(* IEC 61131-3 sources: PLCHoney/Boston Intersection Models/plc_template/webserver/example_st_files, 7 files *)

(* ---- BACNet.st ---- *)
FUNCTION_BLOCK Simulator
  VAR_OUTPUT
    Out : REAL;
  END_VAR
  VAR_INPUT
    MinVal : REAL;
    MaxVal : REAL;
    PeriodSeconds : INT;
  END_VAR
  VAR
    TON0 : TON;
    seconds : INT;
    BaseVal : REAL;
    VarVal : REAL;
  END_VAR

  (* pseudo-random variations *)
  TON0(IN := TRUE, PT := T#3120s);
  IF TON0.Q THEN
    TON0(IN := FALSE);
  END_IF;
  seconds := TIME_TO_INT(TON0.ET);

  BaseVal := (MaxVal + MinVal)/2.0;
  VarVal  := (MaxVal-MinVal)*INT_TO_REAL((seconds MOD PeriodSeconds) - (PeriodSeconds/2))/INT_TO_REAL(PeriodSeconds);

  Out :=  BaseVal + VarVal;
END_FUNCTION_BLOCK

PROGRAM program0
  VAR
    EnergyCounter AT %MD0.2.0 : REAL;
    Temperature AT %ID0.0.0 : REAL;
    Humidity AT %ID0.0.1 : REAL;
  END_VAR
  VAR
    TempSimulation : Simulator;
    HumiditySimulation : Simulator;
  END_VAR
  VAR
    TemperatureSetPoint AT %QD0.1.0 : REAL;
    ControlDisable AT %QX0.4.2 : BOOL;
    Heater AT %IX0.3.0 : BOOL;
    Cooler AT %IX0.3.1 : BOOL;
  END_VAR
  VAR
    ADD3_OUT : REAL;
    GT16_OUT : BOOL;
    AND19_OUT : BOOL;
    LT17_OUT : BOOL;
    AND24_OUT : BOOL;
  END_VAR

  ADD3_OUT := ADD(EnergyCounter, 0.00131);
  EnergyCounter := ADD3_OUT;
  TempSimulation(MinVal := 18.0, MaxVal := 30.0, PeriodSeconds := 120);
  Temperature := TempSimulation.Out;
  HumiditySimulation(MinVal := 55.0, MaxVal := 78.0, PeriodSeconds := 58);
  Humidity := HumiditySimulation.Out;
  GT16_OUT := GT(Temperature, TemperatureSetPoint);
  AND19_OUT := AND(NOT(ControlDisable), GT16_OUT);
  Cooler := AND19_OUT;
  LT17_OUT := LT(Temperature, TemperatureSetPoint);
  AND24_OUT := AND(NOT(ControlDisable), LT17_OUT);
  Heater := AND24_OUT;
END_PROGRAM

CONFIGURATION config

  RESOURCE resource1 ON PLC
    TASK task0(INTERVAL := T#20ms,PRIORITY := 0);
    PROGRAM instance0 WITH task0 : program0;
  END_RESOURCE
END_CONFIGURATION

(* ---- First_Steps.st ---- *)
FUNCTION_BLOCK CounterSFC
  VAR_INPUT
    Reset : BOOL;
  END_VAR
  VAR_OUTPUT
    OUT : INT;
  END_VAR
  VAR
    Cnt : INT;
  END_VAR
  VAR_EXTERNAL CONSTANT
    ResetCounterValue : INT;
  END_VAR

  INITIAL_STEP Start:
  END_STEP

  TRANSITION FROM Start TO ResetCounter
    := Reset;
  END_TRANSITION

  STEP ResetCounter:
    RESETCOUNTER_INLINE1(N);
    RESETCOUNTER_INLINE2(N);
  END_STEP

  ACTION RESETCOUNTER_INLINE1:
    Cnt := ResetCounterValue;
  END_ACTION

  ACTION RESETCOUNTER_INLINE2:
    OUT := Cnt;
  END_ACTION

  TRANSITION FROM ResetCounter TO Start
    := NOT Reset;
  END_TRANSITION

  TRANSITION FROM Start TO Count
    := NOT Reset;
  END_TRANSITION

  STEP Count:
    COUNT_INLINE3(N);
    COUNT_INLINE4(N);
  END_STEP

  ACTION COUNT_INLINE3:
    Cnt := Cnt + 1;
  END_ACTION

  ACTION COUNT_INLINE4:
    OUT := Cnt;
  END_ACTION

  TRANSITION FROM Count TO Start
    := Reset;
  END_TRANSITION

END_FUNCTION_BLOCK

FUNCTION_BLOCK CounterFBD
  VAR_INPUT
    Reset : BOOL;
  END_VAR
  VAR_OUTPUT
    OUT : INT;
  END_VAR
  VAR
    Cnt : INT;
  END_VAR
  VAR_EXTERNAL CONSTANT
    ResetCounterValue : INT;
  END_VAR
  VAR
    ADD4_OUT : INT;
    SEL7_OUT : INT;
  END_VAR

  ADD4_OUT := ADD(1, Cnt);
  SEL7_OUT := SEL(Reset, ADD4_OUT, ResetCounterValue);
  Cnt := SEL7_OUT;
  OUT := Cnt;
END_FUNCTION_BLOCK

FUNCTION_BLOCK CounterIL
  VAR
    Cnt : INT;
  END_VAR
  VAR_INPUT
    Reset : BOOL;
  END_VAR
  VAR_OUTPUT
    OUT : INT;
  END_VAR
  VAR_EXTERNAL CONSTANT
    ResetCounterValue : INT;
  END_VAR

  LD Reset
  JMPC ResetCnt

  (* increment counter *)
  LD Cnt
  ADD 1
  JMP QuitFb

  ResetCnt:
  (* reset counter *)
  LD ResetCounterValue

  QuitFb:
  (* save results *)
  ST Cnt
  ST Out
END_FUNCTION_BLOCK

FUNCTION AverageVal : REAL
  VAR_INPUT
    Cnt1 : INT;
    Cnt2 : INT;
    Cnt3 : INT;
    Cnt4 : INT;
    Cnt5 : INT;
  END_VAR
  VAR
    InputsNumber : REAL := 5.0;
  END_VAR

  AverageVal := INT_TO_REAL(Cnt1+Cnt2+Cnt3+Cnt4+Cnt5)/InputsNumber;
END_FUNCTION

FUNCTION_BLOCK CounterST
  VAR_INPUT
    Reset : BOOL;
  END_VAR
  VAR
    Cnt : INT;
  END_VAR
  VAR_OUTPUT
    OUT : INT;
  END_VAR
  VAR_EXTERNAL CONSTANT
    ResetCounterValue : INT;
  END_VAR

  IF Reset THEN
    Cnt := ResetCounterValue;
  ELSE
    Cnt := Cnt + 1;
  END_IF;

  Out := Cnt;
END_FUNCTION_BLOCK

FUNCTION_BLOCK CounterLD
  VAR_INPUT
    Reset : BOOL;
  END_VAR
  VAR_OUTPUT
    Out : INT;
  END_VAR
  VAR
    Cnt : INT;
  END_VAR
  VAR_EXTERNAL CONSTANT
    ResetCounterValue : INT;
  END_VAR
  VAR
    ADD4_OUT : INT;
    SEL7_OUT : INT;
  END_VAR

  ADD4_OUT := ADD(1, Cnt);
  SEL7_OUT := SEL(Reset, ADD4_OUT, ResetCounterValue);
  Cnt := SEL7_OUT;
  Out := Cnt;
END_FUNCTION_BLOCK

PROGRAM plc_prg
  VAR_INPUT
    Reset : BOOL;
  END_VAR
  VAR_OUTPUT
    Cnt1 : INT;
    Cnt2 : INT;
    Cnt3 : INT;
    Cnt4 : INT;
    Cnt5 : INT;
  END_VAR
  VAR
    CounterST0 : CounterST;
    CounterFBD0 : CounterFBD;
    CounterSFC0 : CounterSFC;
    CounterIL0 : CounterIL;
    CounterLD0 : CounterLD;
    AVCnt : REAL;
    AverageVal17_OUT : REAL;
  END_VAR

  CounterST0(Reset := Reset);
  Cnt1 := CounterST0.OUT;
  AverageVal17_OUT := AverageVal(Cnt1, Cnt2, Cnt3, Cnt4, Cnt5);
  AVCnt := AverageVal17_OUT;
  CounterFBD0(Reset := Reset);
  Cnt2 := CounterFBD0.OUT;
  CounterSFC0(Reset := Reset);
  Cnt3 := CounterSFC0.OUT;
  CounterIL0(Reset := Reset);
  Cnt4 := CounterIL0.OUT;
  CounterLD0(Reset := Reset);
  Cnt5 := CounterLD0.Out;
END_PROGRAM

CONFIGURATION config
  VAR_GLOBAL CONSTANT
    ResetCounterValue : INT := 17;
  END_VAR

  RESOURCE resource1 ON PLC
    TASK plc_task(INTERVAL := T#100ms,PRIORITY := 1);
    PROGRAM plc_task_instance WITH plc_task : plc_prg;
  END_RESOURCE
END_CONFIGURATION

(* ---- modbus.st ---- *)
FUNCTION_BLOCK Generator
  VAR_OUTPUT
    OUT : BOOL;
  END_VAR
  VAR_INPUT
    PON : TIME;
    POFF : TIME;
  END_VAR
  VAR
    T1 : TON;
    T2 : TOF;
  END_VAR

  T1( IN := NOT T2.Q, PT := POFF);
  T2( IN := T1.Q,     PT := PON);
  OUT := T2.Q;
END_FUNCTION_BLOCK

PROGRAM program0
  VAR
    Counter : INT;
    CounterReadBack : INT;
  END_VAR
  VAR
    MasterWriteToReg0 AT %QW0.0.0.0 : INT;
    MasterReadFromReg1 AT %IW0.0.1.0 : INT;
    SlaveHoldReg0 AT %IW0.1.0.0 : WORD;
    SlaveInputReg0 AT %QW0.1.1.0 : WORD;
  END_VAR
  VAR
    CTU0 : CTU;
    Generator0 : Generator;
    R_TRIG1 : R_TRIG;
  END_VAR

  Generator0(PON := T#1s, POFF := T#1s);
  R_TRIG1(CLK := Generator0.OUT);
  CTU0(CU := R_TRIG1.Q, PV := 32767);
  Counter := CTU0.CV;
  MasterWriteToReg0 := Counter;
  CounterReadBack := MasterReadFromReg1;
  SlaveInputReg0 := SlaveHoldReg0;
END_PROGRAM

CONFIGURATION config

  RESOURCE resource1 ON PLC
    TASK task0(INTERVAL := T#20ms,PRIORITY := 0);
    PROGRAM instance0 WITH task0 : program0;
  END_RESOURCE
END_CONFIGURATION

(* ---- canopen_master.st ---- *)
PROGRAM test_main
  VAR
    PLC_OUT AT %QW0.0.2.8193.0 : INT;
    PLC_IN AT %IW0.0.2.8192.0 : INT;
  END_VAR
  VAR
    ADD4_OUT : INT;
  END_VAR

  ADD4_OUT := ADD(1, PLC_IN);
  PLC_OUT := ADD4_OUT;
END_PROGRAM

CONFIGURATION conf

  RESOURCE res ON PLC
    TASK tache(INTERVAL := t#50ms,PRIORITY := 0);
    PROGRAM toto WITH tache : test_main;
  END_RESOURCE
END_CONFIGURATION

(* ---- canopen_slave.st ---- *)
PROGRAM test_main
  VAR
    outvar AT %QW0.0.8192.0 : INT;
    invar AT %IW0.0.8193.0 : INT;
  END_VAR
  VAR
    ADD4_OUT : INT;
  END_VAR

  ADD4_OUT := ADD(1, invar);
  outvar := ADD4_OUT;
END_PROGRAM

CONFIGURATION conf

  RESOURCE res ON PLC
    TASK tache(INTERVAL := T#10ms,PRIORITY := 0);
    PROGRAM toto WITH tache : test_main;
  END_RESOURCE
END_CONFIGURATION

(* ---- genericmake.st ---- *)
PROGRAM program0
  VAR
    LocalVara : INT;
    LocalVarb : INT;
  END_VAR

  LocalVarb := LocalVara;
END_PROGRAM

CONFIGURATION config

  RESOURCE resource1 ON PLC
    TASK Tsk(INTERVAL := T#100ms,PRIORITY := 0);
    PROGRAM Inst WITH Tsk : program0;
  END_RESOURCE
END_CONFIGURATION

(* ---- Hello_World.st ---- *)
PROGRAM Hello_World
  VAR
    my_button AT %IX0.0 : BOOL;
    lamp AT %QX0.0 : BOOL;
  END_VAR
  VAR
    TOF0 : TOF;
  END_VAR

  TOF0(IN := my_button, PT := T#2000ms);
  lamp := TOF0.Q;
END_PROGRAM

CONFIGURATION Config0

  RESOURCE Res0 ON PLC
    TASK task0(INTERVAL := T#20ms,PRIORITY := 0);
    PROGRAM instance0 WITH task0 : Hello_World;
  END_RESOURCE
END_CONFIGURATION
